TYPE "ST_Oee"
VERSION : 0.1
   STRUCT
      "RunMs" : UDInt;
      "DownMs" : UDInt;
      "IdleMs" : UDInt;
      "Availability" : Real;
      "AvailValid" : Bool;
      "Performance" : Real;
      "PerfValid" : Bool;
      "Quality" : Real;
      "QualValid" : Bool;
      "Oee" : Real;
      "OeeValid" : Bool;
      "IdealCycleMs" : UDInt;
   END_STRUCT;
END_TYPE
